(* Logix 5000 project; controller NWGG_Treater_Dayton vendor 1 type 14 code 238 rev 35.11; software revision 35.00; part 3 of 5 *)

ADD_ON_INSTRUCTION SAI_IND_ZeroAdjust   (* revision 1.0, vendor Griffin Hodnett *)
VAR_INPUT
   Start : BOOL; {visible}
END_VAR
VAR_OUTPUT
   Done : BOOL; {access Read Only, visible}
   Error : BOOL; {access Read Only, visible}
   Status : INT; {access Read Only, visible}
END_VAR
VAR_IN_OUT
   MSG_ZeroAdj : MESSAGE; {required}
   MSG_ReadAdjStatus : MESSAGE; {required}
   TmpTrigger : SINT; {required}
   TmpAdjStatus : INT; {required}
END_VAR
VAR
   TON : TIMER[3]; {access None}
   Step : INT; {access None}
   ons : DINT; {access None}
   EnterAdj : BOOL; {access None}
END_VAR

ROUTINE Logic   (* ladder *)
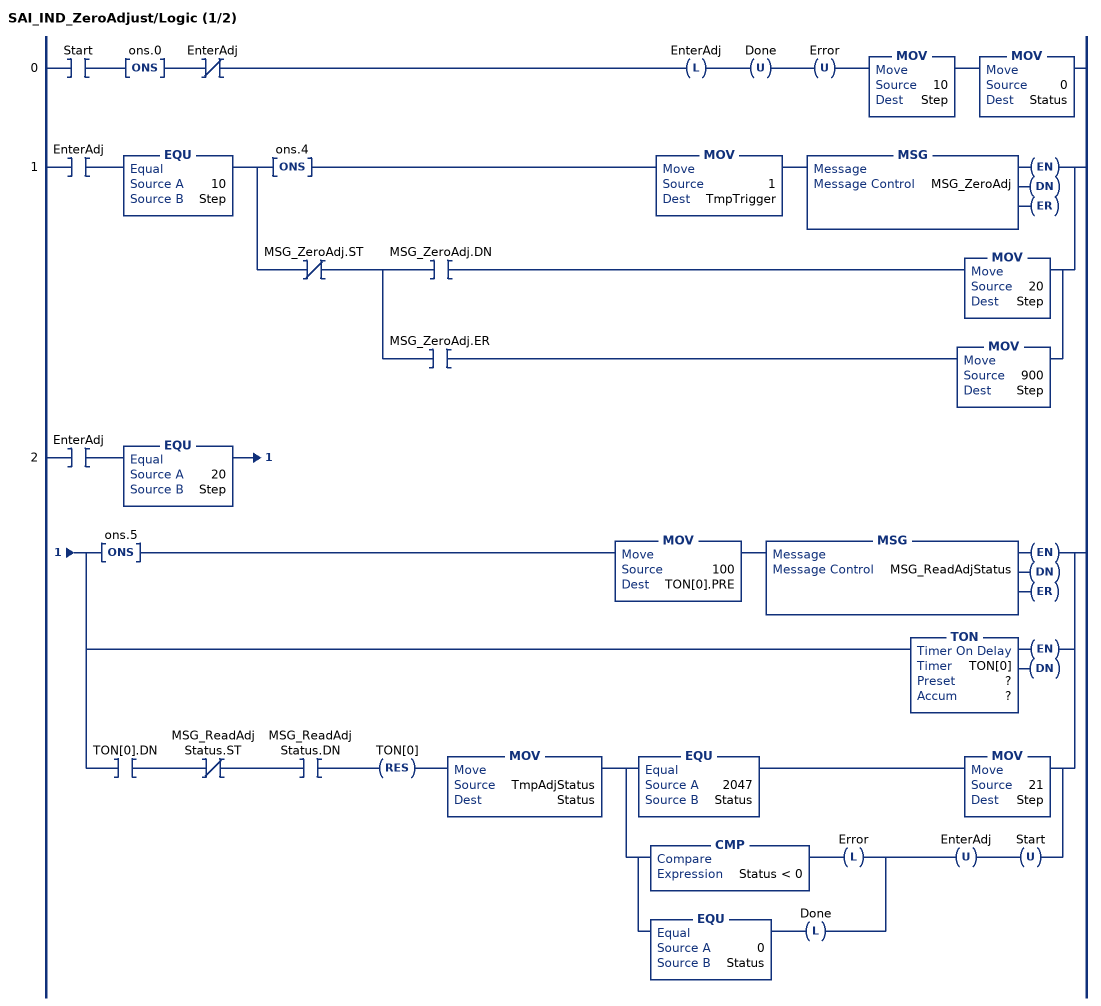
   0: XIC(Start)ONS(ons.0)XIO(EnterAdj)OTL(EnterAdj)OTU(Done)OTU(Error)MOV(10,Step)MOV(0,Status);
   1: XIC(EnterAdj)EQU(10,Step)[ONS(ons.4) MOV(1,TmpTrigger) MSG(MSG_ZeroAdj) ,XIO(MSG_ZeroAdj.ST) [XIC(MSG_ZeroAdj.DN) MOV(20,Step) ,XIC(MSG_ZeroAdj.ER) MOV(900,Step) ] ];
   2: XIC(EnterAdj)EQU(20,Step)[[ONS(ons.5) MOV(100,TON[0].PRE) MSG(MSG_ReadAdjStatus) ,TON(TON[0],?,?) ] ,XIC(TON[0].DN) XIO(MSG_ReadAdjStatus.ST) XIC(MSG_ReadAdjStatus.DN) RES(TON[0]) MOV(TmpAdjStatus,Status) [EQU(2047,Status) MOV(21,Step) ,[CMP(Status < 0) OTL(Error) ,EQU(0,Status) OTL(Done) ] OTU(EnterAdj) OTU(Start) ] ];
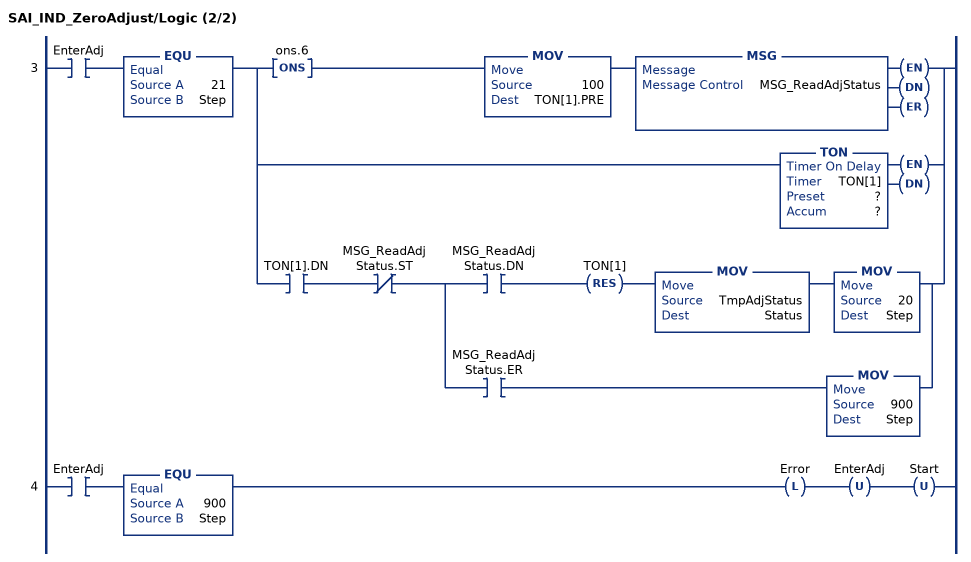
   3: XIC(EnterAdj)EQU(21,Step)[[ONS(ons.6) MOV(100,TON[1].PRE) MSG(MSG_ReadAdjStatus) ,TON(TON[1],?,?) ] ,XIC(TON[1].DN) XIO(MSG_ReadAdjStatus.ST) [XIC(MSG_ReadAdjStatus.DN) RES(TON[1]) MOV(TmpAdjStatus,Status) MOV(20,Step) ,XIC(MSG_ReadAdjStatus.ER) MOV(900,Step) ] ];
   4: XIC(EnterAdj)EQU(900,Step)OTL(Error)OTU(EnterAdj)OTU(Start);
END_ROUTINE
END_ADD_ON_INSTRUCTION

ADD_ON_INSTRUCTION SAI_Scale_Rate   (* revision 1.0, vendor NWGG *)
VAR_INPUT
   UpdateRate : REAL; {access Read Only, required}
END_VAR
VAR_IN_OUT
   Treater_Pump : Treater_Pump; {required}
END_VAR
VAR_INPUT
   Grain_Flow_CWT : REAL; {access None}
END_VAR
VAR
   tmrSecond : TIMER; {access None}
   LastScaleValue : REAL; {access None}
   StartingWeight : REAL; {access None}
   EndingWeight : REAL; {access None}
   LbsRate : REAL; {access None}
   ONS_Output_Bit_1 : BOOL; {access None}
   ONS_Storage_Bit_1 : BOOL; {access None}
END_VAR

ROUTINE Logic   (* ladder *)
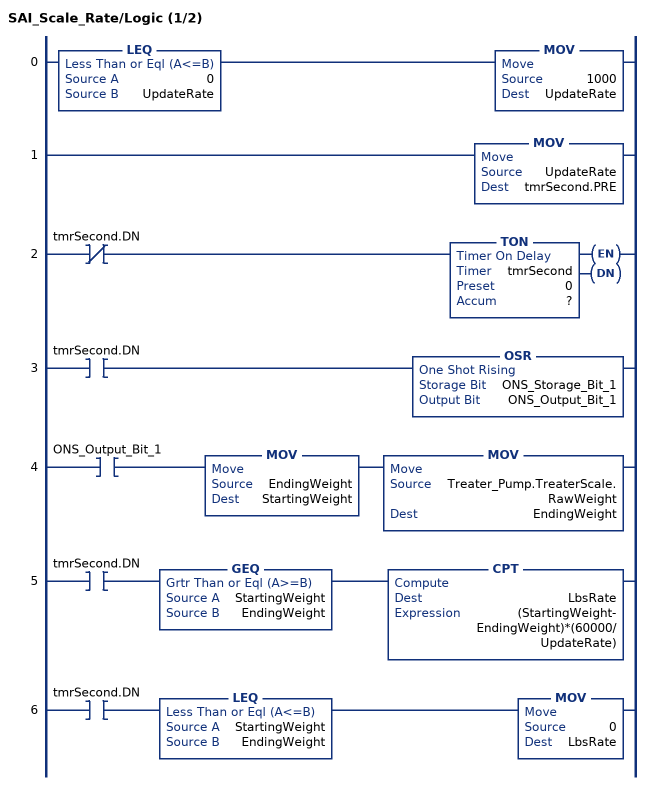
   0: LEQ(0,UpdateRate)MOV(1000,UpdateRate);
   1: MOV(UpdateRate,tmrSecond.PRE);
   2: XIO(tmrSecond.DN)TON(tmrSecond,?,?);
   3: XIC(tmrSecond.DN)OSR(ONS_Storage_Bit_1,ONS_Output_Bit_1);
   4: XIC(ONS_Output_Bit_1)MOV(EndingWeight,StartingWeight)MOV(Treater_Pump.TreaterScale.RawWeight,EndingWeight);
   5: XIC(tmrSecond.DN)GEQ(StartingWeight,EndingWeight)CPT(LbsRate,(StartingWeight-EndingWeight)*(60000/UpdateRate));
   6: XIC(tmrSecond.DN)LEQ(StartingWeight,EndingWeight)MOV(0,LbsRate);
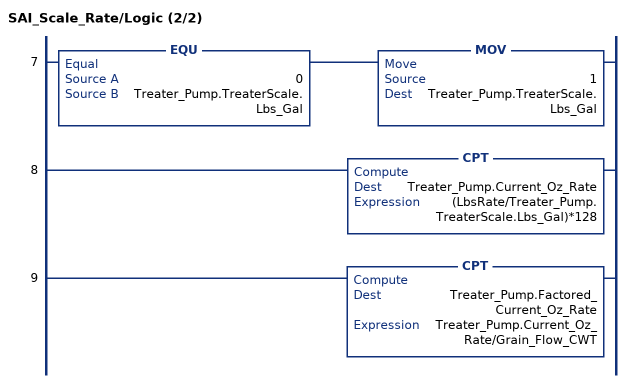
   7: EQU(0,Treater_Pump.TreaterScale.Lbs_Gal)MOV(1,Treater_Pump.TreaterScale.Lbs_Gal);
   8: CPT(Treater_Pump.Current_Oz_Rate,(LbsRate/Treater_Pump.TreaterScale.Lbs_Gal)*128);
   9: CPT(Treater_Pump.Factored_Current_Oz_Rate,Treater_Pump.Current_Oz_Rate/Grain_Flow_CWT);
END_ROUTINE
END_ADD_ON_INSTRUCTION

ADD_ON_INSTRUCTION SAI_Zero_Scale   (* revision 1.0, vendor NWGG *)
VAR_IN_OUT
   MT_ScaleWO : ME:IND360_2BlockW:O:0; {required}
   MT_ScaleWI : ME:IND360_2BlockR:I:0; {required}
   Zero_Scale : BOOL; {required}
END_VAR
VAR
   ZeroCommand : INT; {access Read Only}
   CommandFail : INT; {access Read Only}
   tmrReset : TIMER; {access None}
   ZeroScaleLatch : BOOL; {access None}
END_VAR

ROUTINE Logic   (* ladder *)
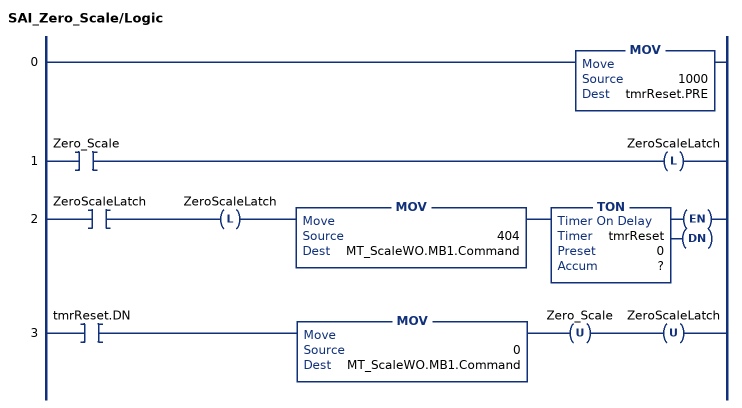
   0: MOV(1000,tmrReset.PRE);
   1: XIC(Zero_Scale)OTL(ZeroScaleLatch);
   2: XIC(ZeroScaleLatch)OTL(ZeroScaleLatch)MOV(404,MT_ScaleWO.MB1.Command)TON(tmrReset,?,?);
   3: XIC(tmrReset.DN)MOV(0,MT_ScaleWO.MB1.Command)OTU(Zero_Scale)OTU(ZeroScaleLatch);
END_ROUTINE
END_ADD_ON_INSTRUCTION

ADD_ON_INSTRUCTION SCP   (* revision 1.2, vendor Rockwell Automation *)
// Scale w/Parameters
// Help:
// Use this instruction to scale data from your analog module and bring it into the limits prescribed by the process variable or another analog module.
// Equations used in calculating a linear relationship:
// Scaled value = (input value - input min.) x rate + scaled minimum
// Rate = (scaled max. - scaled min.) / (input max. - input min.)
VAR_INPUT
   Input : REAL; {required}
   Input_Min : REAL; {required}
   Input_Max : REAL; {required}
   Scaled_Min : REAL; {required}
   Scaled_Max : REAL; {required}
END_VAR
VAR_OUTPUT
   Output : REAL; {access Read Only, required}
END_VAR
VAR
   Rate : REAL;
END_VAR

ROUTINE Logic   (* ladder *)
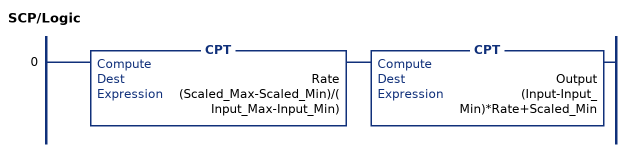
   0: CPT(Rate,(Scaled_Max-Scaled_Min)/(Input_Max-Input_Min))CPT(Output,(Input-Input_Min)*Rate+Scaled_Min);
END_ROUTINE
END_ADD_ON_INSTRUCTION

ADD_ON_INSTRUCTION Water_Pump_Control   (* revision 1.0 *)
VAR_IN_OUT
   Pump_Drive_Out : AB:PowerFlex525V_EENET_Drive:O:0; {required}   // Pump Output
   Pump_Drive_In : AB:PowerFlex525V_EENET_Drive:I:0; {required}   // Pump Input
   Treater_Pump : Treater_Pump; {required}
        .Current_Oz_Rate   // This is the rate adjusted for the Current flow of grain reflected by the muiltliplier
END_VAR
VAR_INPUT
   Grain_Flow_CWT : REAL; {access None, required}
   Pump_Reversed : BOOL; {access Read Only, required}
END_VAR
VAR_IN_OUT
   Values : Analog_Gallon_Values; {required}   // Stored Values
   Analog_Raw_Counts : REAL; {required}
END_VAR
VAR_INPUT
   Start_Treating : BOOL; {access Read Only, required}
   Total_Chemical_Package : REAL; {access Read Only, required}
   Non_Water_Total_Chemical_Package : REAL; {access Read Only, required}
END_VAR
VAR
   Empty_String : STRING; {access None}
   PMC : Pump_Motor_Control; {access None}
   AnalogRate : Analog_Rate; {access None}
   Water_Pump : Analog_Pump_Control; {access None}
END_VAR

ROUTINE Logic   (* ladder *)
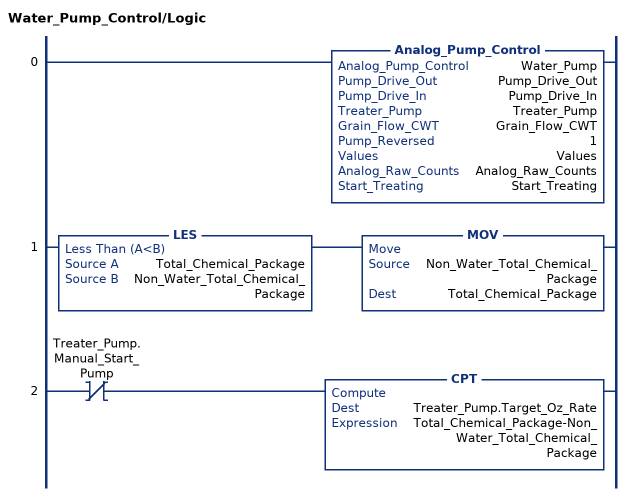
   0: Analog_Pump_Control(Water_Pump,Pump_Drive_Out,Pump_Drive_In,Treater_Pump,Grain_Flow_CWT,1,Values,Analog_Raw_Counts,Start_Treating);
   1: LES(Total_Chemical_Package,Non_Water_Total_Chemical_Package)MOV(Non_Water_Total_Chemical_Package,Total_Chemical_Package);
   2: XIO(Treater_Pump.Manual_Start_Pump)CPT(Treater_Pump.Target_Oz_Rate,Total_Chemical_Package-Non_Water_Total_Chemical_Package);
END_ROUTINE
END_ADD_ON_INSTRUCTION

VAR_GLOBAL   (* controller tags *)
   Auto_Start_Treater : BOOL;
   Check_For_Flush : BOOL := 1;
   Chemicals_Required : BOOL;
   Clear_Treater_Fault : BOOL := 1;
   Color_Index : INT;
   Colors : Color[10];
   Current_Color : Color;   // Current Color Being Used
   Current_Rate : REAL := 10.5;
   Current_Treater_Pump : Active_Pump_Values[6];
   Current_Treater_Speed_Percent : REAL;
   Default_Speed_Factor : REAL;   // The default factor used for pump rpm
   Edit_Color : Color;
   Edit_Color_Idx : DINT := 2;
   Edit_Idx : INT;
   Grain_Rate_CWT : REAL := 17.12;
   IDX : DINT := 22;
   K_Valve_ACK : BOOL;
   LinearityRange_1 : INT;
   Long_Belt_Amps : REAL := 0.032609403;
   Long_Belt_SCP : SCP;
   Manual_Start_Treater : BOOL;
   Manual_Stop_Pumps : BOOL;
   Non_Water_Total_Chemical_Package : REAL;
   Non_Water_Treatment_Package : REAL := 14.209999;
   PumpParams : PumpParameters[32];
   RatedCapacity_1 : REAL;
   RatedOutput_1 : REAL;
   RatePid : PID[32];
   SAIZeroScale : SAI_Zero_Scale[30]; {access Read Only}
   SaveEdit : BOOL;
   ScaleUnit_1 : SINT;
   Start_Treater : BOOL;
   Start_Treating : BOOL;
   Stop_Treater : BOOL;
   Stop_Treating : BOOL;
   TestLong : DINT;   // Test Dint
   TmpAdjStatus_1 : INT;
   TmpAdjTrigger_1 : SINT;
   TmpCalFreeTrigger_1 : INT;
   TmpCapacity_1 : REAL;
   TmpIncrement_1 : REAL;
   TmpSpanAdjWeight_1 : REAL;
   tmrStartTreat : TIMER;
   tmrStopTreat : TIMER;
   tmrZtest : TIMER; {access Read Only}
   Total_Chemical_Package : REAL := 18.0;
   Total_CWT_Min : DINT; {access Read Only}
   Treater_Pump : Treater_Pump[50];
        [5].Target_Oz_Rate   // Mineral Oil lbs/min Called For
        [1].Target_Oz_Rate   // Blue The lbs/min called For
        [3].Start_Pump   // Yellow Bit To Start The Pump
        [0]   // Water
        [1].Active_Treatment   // Water Used In Batch
        [2].Start_Pump   // Red Bit To Start The Pump
        [22].Manual_Start_Pump   // Water Manual Start Pump
        [2].Target_Oz_Rate   // Red lbs / Min Called For
        [3].Manual_Start_Pump   // Yellow Manual Pump Start
        [3].Target_Oz_Rate   // Yellow lbs/ min Called For
        [1].Manual_Start_Pump   // Blue Manual Start Pump
        [2]   // Red
        [2].Manual_Start_Pump   // Red Manual Pump Start
        [3]   // Yellow
        [4]   // Mineral
        [1]   // Blue
        [5]   // Rinseate
        [22].Target_Oz_Rate   // Water pounds/min called for
        [5].Active_Treatment   // Mineral Oil Used In Batch
   Treater_Pump_Fault : BOOL;
   Treater_Running : BOOL;
   Treater_Speed_Percent : REAL := 1.0;
   Treatment_Products : Treater_Product[100];   // The List Of Treater Products Used
   Use_Mineral_Oil : BOOL;
   Use_Oil_In_Treat : BOOL;
   UseScales : BOOL;
   Water : Analog_Gallon_Values;
   Water_Control : Water_Pump_Control;
   Water_Pump : Analog_Pump_Control;
   WriteAdjustSettings_Capacity_1 : REAL;
   WriteAdjustSettings_Increment_1 : REAL;
END_VAR

PROGRAM ColorBlending   (* main routine Blending *)
VAR
   BlendColorCount : INT := 1;
   Blue_Pump : Treater_Pump;
   BlueRate : REAL;
   ColorCountIdx : INT;
   ColorIndexChanged : BOOL;
   CountIdx : DINT := 10;
   ctrColorIdx : COUNTER;
   ctrIndex : COUNTER;
   CurColorIdx : INT;
   IDX : INT := 5;
   Inactive_Color : BOOL;
   Initialize : BOOL;
   NewColorIdx : INT;
   NextColor : BOOL;
   NextColorSet : BOOL;
   No_Color : BOOL := 1;
   Pause : BOOL := 1;
   PolymerRate : REAL := 10.25;
   PumpDelay : DINT;
   RedRate : REAL := 20.5;
   ReverseDuration : DINT;
   ReverseONS : BOOL := 1;
   ReverseRate : REAL := 20.0;
   ReverseStart : BOOL;
   SetColorIndex : BOOL;
   SetReverseRate : BOOL;
   Start_Color : BOOL;
   TestBit : BOOL;
   testReal : REAL;
   TestReverse : BOOL;
   tmrDelay : TIMER;
   tmrDuration : TIMER;
   tmrReverse : TIMER;
   Total_Oz_Min : DINT := 41;
   WhiteRate : REAL;
   YellowRate : REAL;
END_VAR

ROUTINE Blending   (* ladder *)
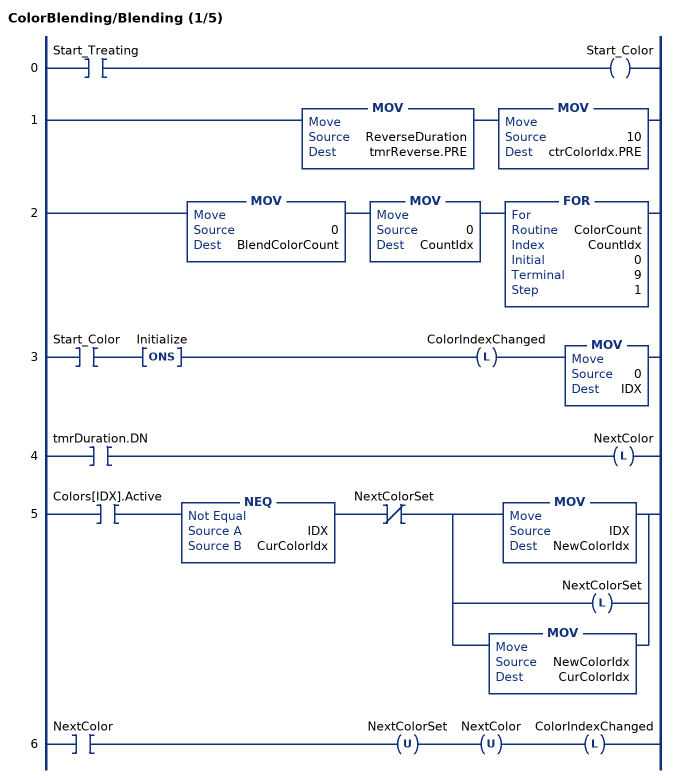
   0: XIC(Start_Treating)OTE(Start_Color);
   1: MOV(ReverseDuration,tmrReverse.PRE)MOV(10,ctrColorIdx.PRE);
   2: MOV(0,BlendColorCount)MOV(0,CountIdx)FOR(ColorCount,CountIdx,0,9,1);
   3: XIC(Start_Color)ONS(Initialize)OTL(ColorIndexChanged)MOV(0,IDX);
   4: XIC(tmrDuration.DN)OTL(NextColor);
   5: XIC(Colors[IDX].Active)NEQ(IDX,CurColorIdx)XIO(NextColorSet)[MOV(IDX,NewColorIdx) ,OTL(NextColorSet) ,MOV(NewColorIdx,CurColorIdx) ];
   6: XIC(NextColor)OTU(NextColorSet)OTU(NextColor)OTL(ColorIndexChanged);
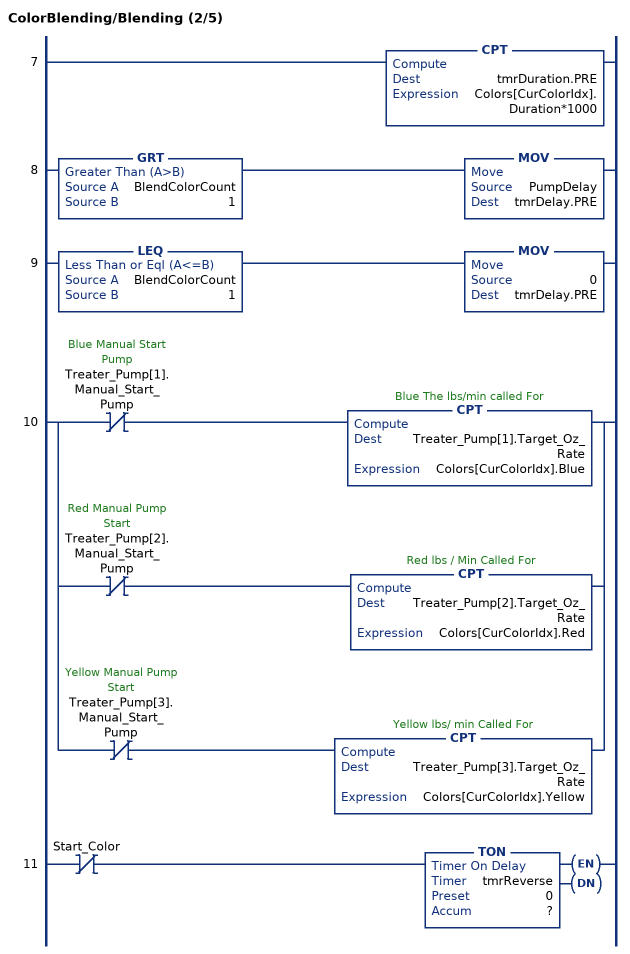
   7: CPT(tmrDuration.PRE,Colors[CurColorIdx].Duration*1000);
   8: GRT(BlendColorCount,1)MOV(PumpDelay,tmrDelay.PRE);
   9: LEQ(BlendColorCount,1)MOV(0,tmrDelay.PRE);
   10: [XIO(Treater_Pump[1].Manual_Start_Pump) CPT(Treater_Pump[1].Target_Oz_Rate,Colors[CurColorIdx].Blue) ,XIO(Treater_Pump[2].Manual_Start_Pump) CPT(Treater_Pump[2].Target_Oz_Rate,Colors[CurColorIdx].Red) ,XIO(Treater_Pump[3].Manual_Start_Pump) CPT(Treater_Pump[3].Target_Oz_Rate,Colors[CurColorIdx].Yellow) ];
   11: XIO(Start_Color)TON(tmrReverse,?,?);
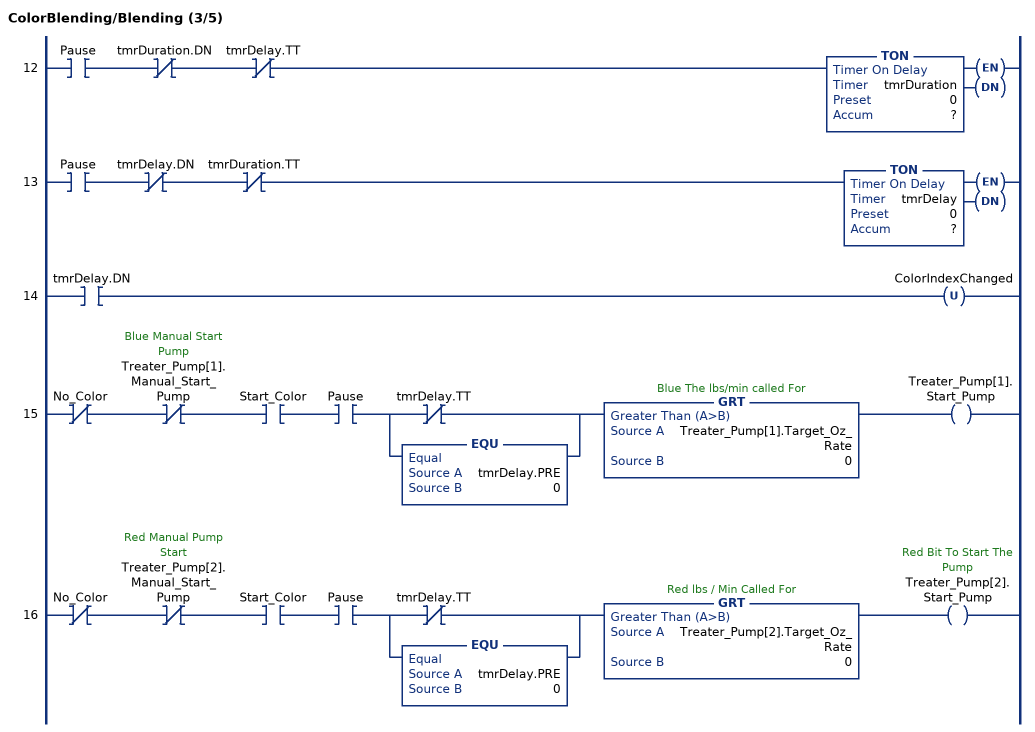
   12: XIC(Pause)XIO(tmrDuration.DN)XIO(tmrDelay.TT)TON(tmrDuration,?,?);
   13: XIC(Pause)XIO(tmrDelay.DN)XIO(tmrDuration.TT)TON(tmrDelay,?,?);
   14: XIC(tmrDelay.DN)OTU(ColorIndexChanged);
   15: XIO(No_Color)XIO(Treater_Pump[1].Manual_Start_Pump)XIC(Start_Color)XIC(Pause)[XIO(tmrDelay.TT) ,EQU(tmrDelay.PRE,0) ]GRT(Treater_Pump[1].Target_Oz_Rate,0)OTE(Treater_Pump[1].Start_Pump);
   16: XIO(No_Color)XIO(Treater_Pump[2].Manual_Start_Pump)XIC(Start_Color)XIC(Pause)[XIO(tmrDelay.TT) ,EQU(tmrDelay.PRE,0) ]GRT(Treater_Pump[2].Target_Oz_Rate,0)OTE(Treater_Pump[2].Start_Pump);
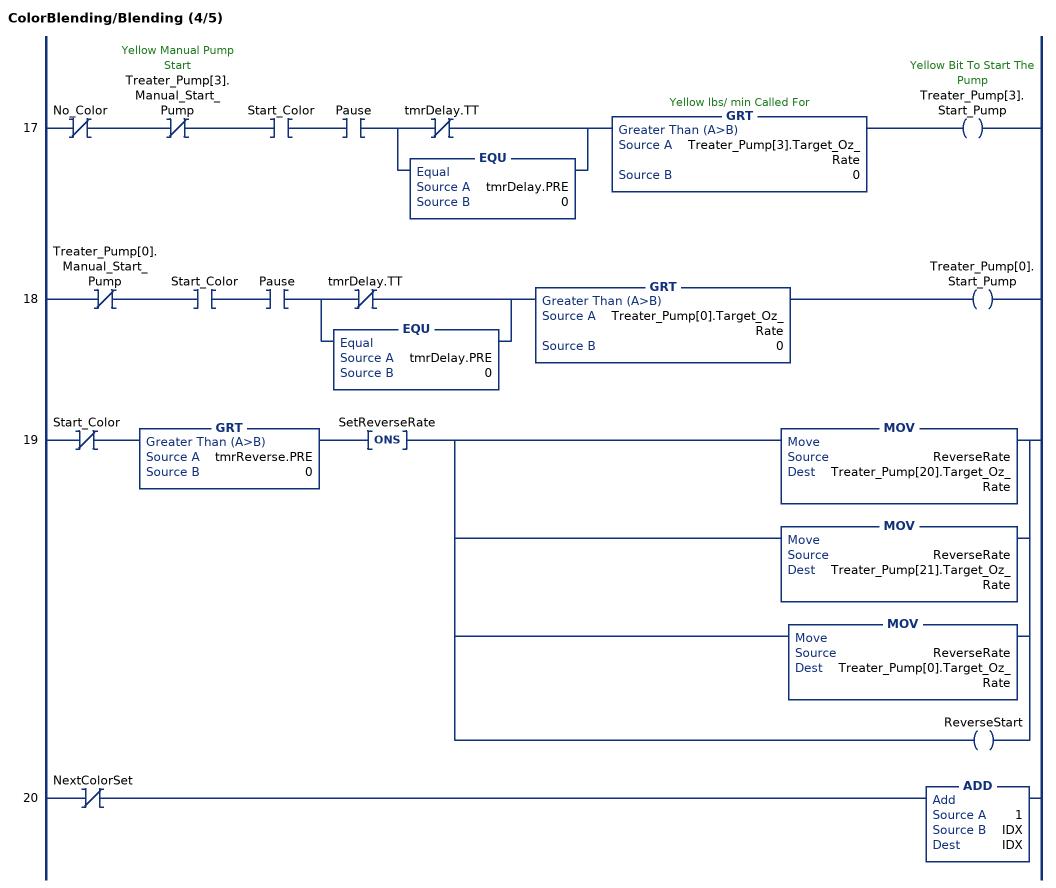
   17: XIO(No_Color)XIO(Treater_Pump[3].Manual_Start_Pump)XIC(Start_Color)XIC(Pause)[XIO(tmrDelay.TT) ,EQU(tmrDelay.PRE,0) ]GRT(Treater_Pump[3].Target_Oz_Rate,0)OTE(Treater_Pump[3].Start_Pump);
   18: XIO(Treater_Pump[0].Manual_Start_Pump)XIC(Start_Color)XIC(Pause)[XIO(tmrDelay.TT) ,EQU(tmrDelay.PRE,0) ]GRT(Treater_Pump[0].Target_Oz_Rate,0)OTE(Treater_Pump[0].Start_Pump);
   19: XIO(Start_Color)GRT(tmrReverse.PRE,0)ONS(SetReverseRate)[MOV(ReverseRate,Treater_Pump[20].Target_Oz_Rate) ,MOV(ReverseRate,Treater_Pump[21].Target_Oz_Rate) ,MOV(ReverseRate,Treater_Pump[0].Target_Oz_Rate) ,OTE(ReverseStart) ];
   20: XIO(NextColorSet)ADD(1,IDX,IDX);
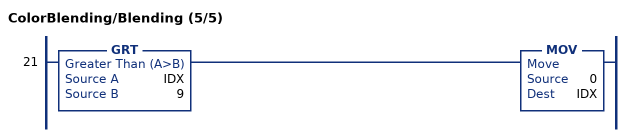
   21: GRT(IDX,9)MOV(0,IDX);
END_ROUTINE

ROUTINE ColorCount   (* ladder *)
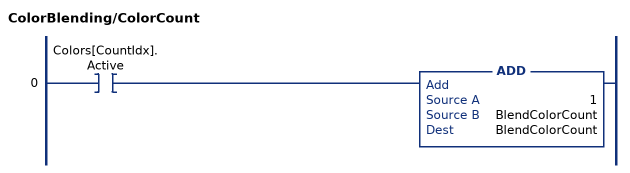
   0: XIC(Colors[CountIdx].Active)ADD(1,BlendColorCount,BlendColorCount);
END_ROUTINE
END_PROGRAM

PROGRAM MainProgram   (* main routine MainRoutine *)
VAR
   ColorPumps : ColorBlending;
   Pump_Product_Description : STRING[30];
   SAI_CheckAlive : SAI_CheckAlive;
   SAI_IND_CalFree : SAI_IND_CalFree;
   SAI_IND_ReadAdjustSettings : SAI_IND_ReadAdjustSettings;
   SAI_IND_SpanAdjust : SAI_IND_SpanAdjust;
   SAI_IND_WeightProc : SAI_IND_WeightProc;
   SAI_IND_WriteAdjustSettings : SAI_IND_WriteAdjustSettings;
   SAI_IND_ZeroAdjust : SAI_IND_ZeroAdjust;
   SAITruckScaleRate : SAI_Scale_Rate; {access Read Only}
   tmrSecond : TIMER; {access Read Only}
   TONR_01 : FBD_TIMER;
END_VAR

ROUTINE Const   (* ladder *)
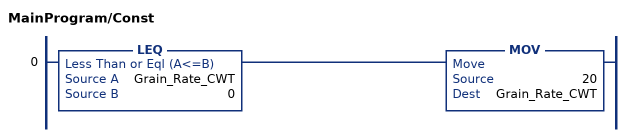
   0: LEQ(Grain_Rate_CWT,0)MOV(20,Grain_Rate_CWT);
END_ROUTINE

ROUTINE MainRoutine   (* ladder *)
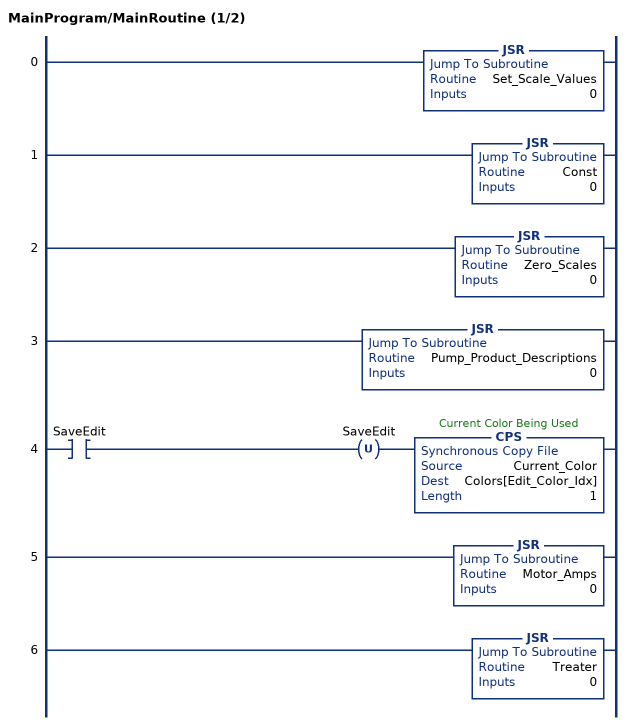
   0: JSR(Set_Scale_Values,0);
   1: JSR(Const,0);
   2: JSR(Zero_Scales,0);
   3: JSR(Pump_Product_Descriptions,0);
   4: XIC(SaveEdit)OTU(SaveEdit)CPS(Current_Color,Colors[Edit_Color_Idx],1);
   5: JSR(Motor_Amps,0);
   6: JSR(Treater,0);
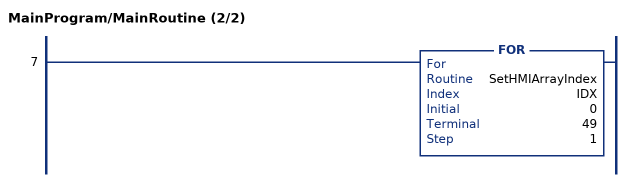
   7: FOR(SetHMIArrayIndex,IDX,0,49,1);
END_ROUTINE

ROUTINE Motor_Amps   (* ladder *)
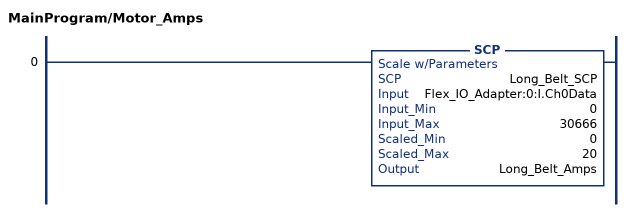
   0: SCP(Long_Belt_SCP,Flex_IO_Adapter:0:I.Ch0Data,0,30666,0,20,Long_Belt_Amps);
END_ROUTINE

ROUTINE Pump_Product_Descriptions   (* ladder *)
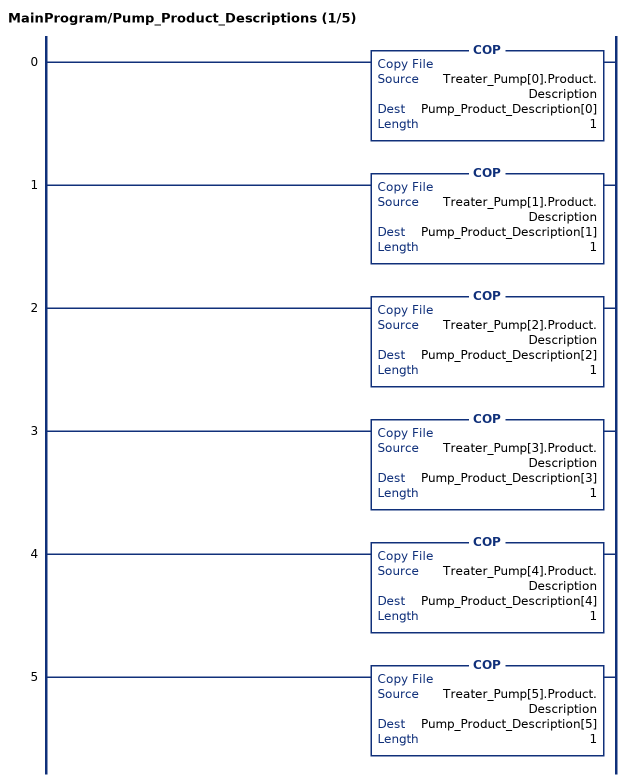
   0: COP(Treater_Pump[0].Product.Description,Pump_Product_Description[0],1);
   1: COP(Treater_Pump[1].Product.Description,Pump_Product_Description[1],1);
   2: COP(Treater_Pump[2].Product.Description,Pump_Product_Description[2],1);
   3: COP(Treater_Pump[3].Product.Description,Pump_Product_Description[3],1);
   4: COP(Treater_Pump[4].Product.Description,Pump_Product_Description[4],1);
   5: COP(Treater_Pump[5].Product.Description,Pump_Product_Description[5],1);
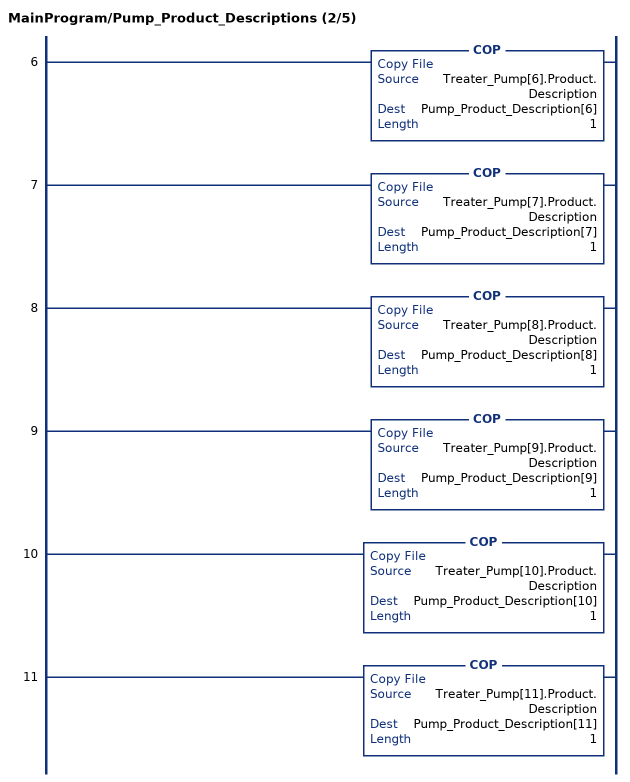
   6: COP(Treater_Pump[6].Product.Description,Pump_Product_Description[6],1);
   7: COP(Treater_Pump[7].Product.Description,Pump_Product_Description[7],1);
   8: COP(Treater_Pump[8].Product.Description,Pump_Product_Description[8],1);
   9: COP(Treater_Pump[9].Product.Description,Pump_Product_Description[9],1);
   10: COP(Treater_Pump[10].Product.Description,Pump_Product_Description[10],1);
   11: COP(Treater_Pump[11].Product.Description,Pump_Product_Description[11],1);
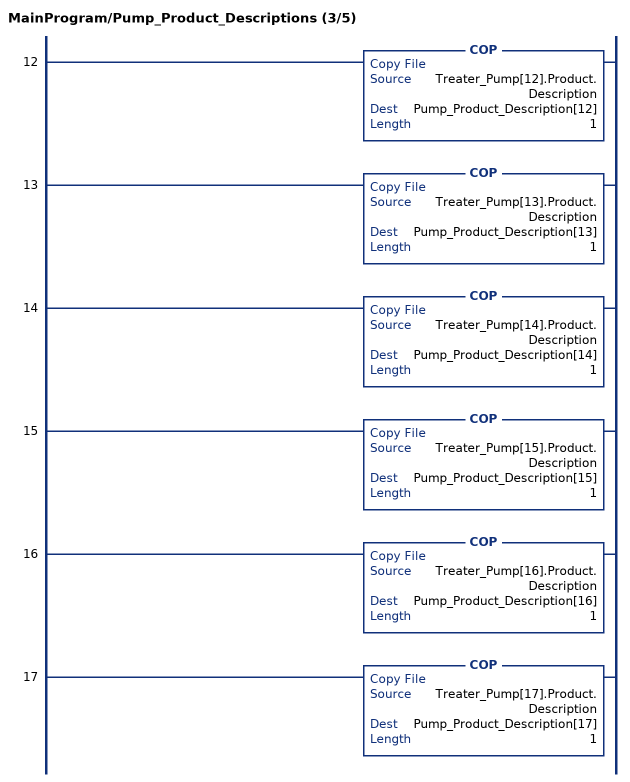
   12: COP(Treater_Pump[12].Product.Description,Pump_Product_Description[12],1);
   13: COP(Treater_Pump[13].Product.Description,Pump_Product_Description[13],1);
   14: COP(Treater_Pump[14].Product.Description,Pump_Product_Description[14],1);
   15: COP(Treater_Pump[15].Product.Description,Pump_Product_Description[15],1);
   16: COP(Treater_Pump[16].Product.Description,Pump_Product_Description[16],1);
   17: COP(Treater_Pump[17].Product.Description,Pump_Product_Description[17],1);
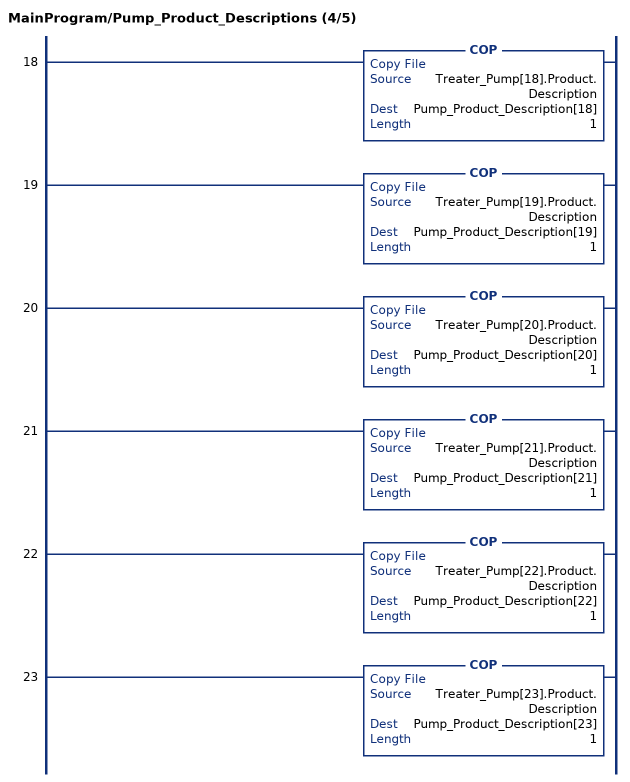
   18: COP(Treater_Pump[18].Product.Description,Pump_Product_Description[18],1);
   19: COP(Treater_Pump[19].Product.Description,Pump_Product_Description[19],1);
   20: COP(Treater_Pump[20].Product.Description,Pump_Product_Description[20],1);
   21: COP(Treater_Pump[21].Product.Description,Pump_Product_Description[21],1);
   22: COP(Treater_Pump[22].Product.Description,Pump_Product_Description[22],1);
   23: COP(Treater_Pump[23].Product.Description,Pump_Product_Description[23],1);
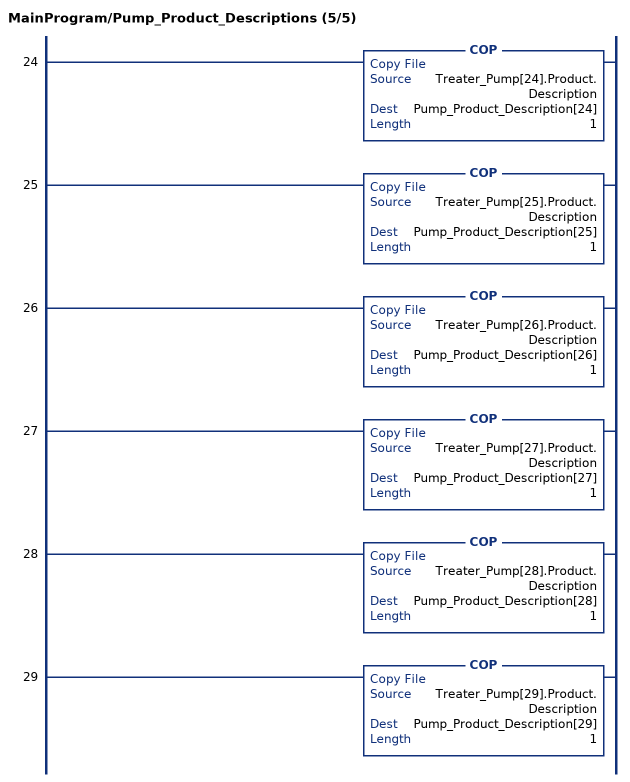
   24: COP(Treater_Pump[24].Product.Description,Pump_Product_Description[24],1);
   25: COP(Treater_Pump[25].Product.Description,Pump_Product_Description[25],1);
   26: COP(Treater_Pump[26].Product.Description,Pump_Product_Description[26],1);
   27: COP(Treater_Pump[27].Product.Description,Pump_Product_Description[27],1);
   28: COP(Treater_Pump[28].Product.Description,Pump_Product_Description[28],1);
   29: COP(Treater_Pump[29].Product.Description,Pump_Product_Description[29],1);
END_ROUTINE
